(* IEC 61131-3 sources: s7-to-codesys/src/POUs/S7Compat/F_S7EnoAddDint, 1 file *)

(* ---- F_S7EnoAddDint.decl.st ---- *)
// Назначение: ENO инструкции S7 ADD (DInt) для кода, сконвертированного s7conv из LAD/FBD:
//             TRUE, если сумма помещается в DINT (-2147483648…2147483647), FALSE при
//             переполнении. У S7 ENO = EN AND NOT переполнение (справочник LAD S7-300/400, прил. C.1),
//             в CODESYS ENO = EN. Результат операции вычисляет вызывающий код; функцию вызывают до записи
//             результата.
// Автор:      kr0nsch
// Версия:     1.1.0
// Документ:   docs/MAPPING_LADFBD.md, правило lad.eno_error
FUNCTION F_S7EnoAddDint : BOOL
VAR_INPUT
    diIn1 : DINT;    // первое слагаемое (IN1)
    diIn2 : DINT;    // второе слагаемое (IN2)
END_VAR
VAR
    liResult : LINT;  // точный результат в LINT
END_VAR
VAR CONSTANT
    DINT_MIN : LINT := -2147483648;   // нижняя граница DINT
    DINT_MAX : LINT := 2147483647;   // верхняя граница DINT
END_VAR
